// TIA Portal V15.1 export
// export: Created 2026-11-01T00:00:00Z, ExportSetting WithDefaults
TagTable "LCP01"
  BR01_TeA : Int  (PLC tag BR01_DB.TeA, HMI_Connection_1, 1 s)
  BR01_TeB : Int  (PLC tag BR01_DB.TeB, HMI_Connection_1, 1 s)
  BR01_Tmax : Int  (PLC tag BR01_DB.Tmax, HMI_Connection_1, 1 s)
  BR01_TcOkA : Bool  (PLC tag BR01_DB.TcOkA, HMI_Connection_1, 1 s)
  BR01_TcOkB : Bool  (PLC tag BR01_DB.TcOkB, HMI_Connection_1, 1 s)
  BR01_TcOk : Bool  (PLC tag BR01_DB.TcOk, HMI_Connection_1, 1 s)
  BR01_State : Int  (PLC tag BR01_DB.State, HMI_Connection_1, 1 s)
  BR01_Enabled : Bool  (PLC tag BR01_DB.Enabled, HMI_Connection_1, 1 s)
  BR01_HeatReq : Bool  (PLC tag BR01_DB.HeatReq, HMI_Connection_1, 1 s)
  BR01_Stage2 : Bool  (PLC tag BR01_DB.Stage2, HMI_Connection_1, 1 s)
  BR01_RunFb : Bool  (PLC tag BR01_DB.RunFb, HMI_Connection_1, 1 s)
  BR01_Lockout : Bool  (PLC tag BR01_DB.Lockout, HMI_Connection_1, 1 s)
  BR01_LevelOK : Bool  (PLC tag BR01_DB.LevelOK, HMI_Connection_1, 1 s)
  BR01_Auto : Bool  (PLC tag BR01_DB.Auto, HMI_Connection_1, 1 s)
  BR01_PwrUpDone : Bool  (PLC tag BR01_DB.PwrUpDone, HMI_Connection_1, 1 s)
  BR01_SP_Act : Int  (PLC tag BR01_DB.SP_Act, HMI_Connection_1, 1 s)
  BR01_TOn : Int  (PLC tag BR01_DB.TOn, HMI_Connection_1, 1 s)
  BR01_TStg : Int  (PLC tag BR01_DB.TStg, HMI_Connection_1, 1 s)
  BR01_TStgOff : Int  (PLC tag BR01_DB.TStgOff, HMI_Connection_1, 1 s)
  BR01_ParPending : Bool  (PLC tag BR01_DB.ParPending, HMI_Connection_1, 1 s)
  BR01_F_EStop : Bool  (PLC tag BR01_DB.F_EStop, HMI_Connection_1, 1 s)
  BR01_F_TC : Bool  (PLC tag BR01_DB.F_TC, HMI_Connection_1, 1 s)
  BR01_F_Lockout : Bool  (PLC tag BR01_DB.F_Lockout, HMI_Connection_1, 1 s)
  BR01_F_NoStart : Bool  (PLC tag BR01_DB.F_NoStart, HMI_Connection_1, 1 s)
  BR01_F_RunLost : Bool  (PLC tag BR01_DB.F_RunLost, HMI_Connection_1, 1 s)
  BR01_F_RunWrong : Bool  (PLC tag BR01_DB.F_RunWrong, HMI_Connection_1, 1 s)
  BR01_Pause24 : Bool  (PLC tag BR01_DB.Pause24, HMI_Connection_1, 1 s)
  BR02_TeA : Int  (PLC tag BR02_DB.TeA, HMI_Connection_1, 1 s)
  BR02_TeB : Int  (PLC tag BR02_DB.TeB, HMI_Connection_1, 1 s)
  BR02_Tmax : Int  (PLC tag BR02_DB.Tmax, HMI_Connection_1, 1 s)
  BR02_TcOkA : Bool  (PLC tag BR02_DB.TcOkA, HMI_Connection_1, 1 s)
  BR02_TcOkB : Bool  (PLC tag BR02_DB.TcOkB, HMI_Connection_1, 1 s)
  BR02_TcOk : Bool  (PLC tag BR02_DB.TcOk, HMI_Connection_1, 1 s)
  BR02_State : Int  (PLC tag BR02_DB.State, HMI_Connection_1, 1 s)
  BR02_Enabled : Bool  (PLC tag BR02_DB.Enabled, HMI_Connection_1, 1 s)
  BR02_HeatReq : Bool  (PLC tag BR02_DB.HeatReq, HMI_Connection_1, 1 s)
  BR02_Stage2 : Bool  (PLC tag BR02_DB.Stage2, HMI_Connection_1, 1 s)
  BR02_RunFb : Bool  (PLC tag BR02_DB.RunFb, HMI_Connection_1, 1 s)
  BR02_Lockout : Bool  (PLC tag BR02_DB.Lockout, HMI_Connection_1, 1 s)
  BR02_LevelOK : Bool  (PLC tag BR02_DB.LevelOK, HMI_Connection_1, 1 s)
  BR02_Auto : Bool  (PLC tag BR02_DB.Auto, HMI_Connection_1, 1 s)
  BR02_PwrUpDone : Bool  (PLC tag BR02_DB.PwrUpDone, HMI_Connection_1, 1 s)
  BR02_SP_Act : Int  (PLC tag BR02_DB.SP_Act, HMI_Connection_1, 1 s)
  BR02_TOn : Int  (PLC tag BR02_DB.TOn, HMI_Connection_1, 1 s)
  BR02_TStg : Int  (PLC tag BR02_DB.TStg, HMI_Connection_1, 1 s)
  BR02_TStgOff : Int  (PLC tag BR02_DB.TStgOff, HMI_Connection_1, 1 s)
  BR02_ParPending : Bool  (PLC tag BR02_DB.ParPending, HMI_Connection_1, 1 s)
  BR02_F_EStop : Bool  (PLC tag BR02_DB.F_EStop, HMI_Connection_1, 1 s)
  BR02_F_TC : Bool  (PLC tag BR02_DB.F_TC, HMI_Connection_1, 1 s)
  BR02_F_Lockout : Bool  (PLC tag BR02_DB.F_Lockout, HMI_Connection_1, 1 s)
  BR02_F_NoStart : Bool  (PLC tag BR02_DB.F_NoStart, HMI_Connection_1, 1 s)
  BR02_F_RunLost : Bool  (PLC tag BR02_DB.F_RunLost, HMI_Connection_1, 1 s)
  BR02_F_RunWrong : Bool  (PLC tag BR02_DB.F_RunWrong, HMI_Connection_1, 1 s)
  BR02_Fuel : Bool  (PLC tag BR02_DB.Fuel, HMI_Connection_1, 1 s)
  Scrub_PSH : Bool  (PLC tag Scrubber_DB.PSH, HMI_Connection_1, 1 s)
  Scrub_LSH : Bool  (PLC tag Scrubber_DB.LSH, HMI_Connection_1, 1 s)
  Scrub_LSHH : Bool  (PLC tag Scrubber_DB.LSHH, HMI_Connection_1, 1 s)
  Scrub_Tripped : Bool  (PLC tag Scrubber_DB.Tripped, HMI_Connection_1, 1 s)
  Scrub_ValvesNormal : Bool  (PLC tag Scrubber_DB.ValvesNormal, HMI_Connection_1, 1 s)
  Scrub_Cause_EStop : Bool  (PLC tag Scrubber_DB.Cause_EStop, HMI_Connection_1, 1 s)
  Scrub_Cause_PSH : Bool  (PLC tag Scrubber_DB.Cause_PSH, HMI_Connection_1, 1 s)
  Scrub_Cause_LSHH : Bool  (PLC tag Scrubber_DB.Cause_LSHH, HMI_Connection_1, 1 s)
  Scrub_Cause_PwrUp : Bool  (PLC tag Scrubber_DB.Cause_PwrUp, HMI_Connection_1, 1 s)
  Scrub_FirstOut : Int  (PLC tag Scrubber_DB.FirstOut, HMI_Connection_1, 1 s)
  Scrub_FlareCmd : Bool  (PLC tag Scrubber_DB.FlareCmd, HMI_Connection_1, 1 s)
  Scrub_DrainCmd : Bool  (PLC tag Scrubber_DB.DrainCmd, HMI_Connection_1, 1 s)
  Scrub_SuctionCmd : Bool  (PLC tag Scrubber_DB.SuctionCmd, HMI_Connection_1, 1 s)
  Scrub_F_DrainTO : Bool  (PLC tag Scrubber_DB.F_DrainTO, HMI_Connection_1, 1 s)
  Scrub_F_LshFault : Bool  (PLC tag Scrubber_DB.F_LshFault, HMI_Connection_1, 1 s)
  Par_SP : Int  (PLC tag Par.SP, HMI_Connection_1, 1 s)
  Par_HYST : Int  (PLC tag Par.HYST, HMI_Connection_1, 1 s)
  Par_STG : Int  (PLC tag Par.STG, HMI_Connection_1, 1 s)
  Par_TStart : Time  (PLC tag Par.TStart, HMI_Connection_1, 1 s)
  Par_TDrnOn : Time  (PLC tag Par.TDrnOn, HMI_Connection_1, 1 s)
  Par_TDrnOff : Time  (PLC tag Par.TDrnOff, HMI_Connection_1, 1 s)
  Par_TDrnMax : Time  (PLC tag Par.TDrnMax, HMI_Connection_1, 1 s)
  Par_SP_V : Int  (PLC tag Par.SP_V, HMI_Connection_1, 1 s)
  Par_HYST_V : Int  (PLC tag Par.HYST_V, HMI_Connection_1, 1 s)
  Par_STG_V : Int  (PLC tag Par.STG_V, HMI_Connection_1, 1 s)
  Par_TStart_V : Time  (PLC tag Par.TStart_V, HMI_Connection_1, 1 s)
  Par_TDrnOn_V : Time  (PLC tag Par.TDrnOn_V, HMI_Connection_1, 1 s)
  Par_TDrnOff_V : Time  (PLC tag Par.TDrnOff_V, HMI_Connection_1, 1 s)
  Par_TDrnMax_V : Time  (PLC tag Par.TDrnMax_V, HMI_Connection_1, 1 s)
  Sys_EStopOK : Bool  (PLC tag Sys.EStopOK, HMI_Connection_1, 1 s)
  Sys_Alm_EStop : Bool  (PLC tag Sys.Alm_EStop, HMI_Connection_1, 1 s)
  Sys_Alm_ParRejected : Bool  (PLC tag Sys.Alm_ParRejected, HMI_Connection_1, 1 s)
  Alm_Common : Word  (PLC tag HmiAlm.Common, HMI_Connection_1, 1 s)
  Alm_BR01 : Word  (PLC tag HmiAlm.BR01, HMI_Connection_1, 1 s)
  Alm_BR02 : Word  (PLC tag HmiAlm.BR02, HMI_Connection_1, 1 s)
